Fanuc KAREL source: KX00016.KL

PROGRAM KX00016
%NOLOCKGROUP
VAR
  I: INTEGER
  J: INTEGER
  B: BOOLEAN
  F: FILE
  S: STRING[80]
  P: XYZWPR
BEGIN
  ENABLE CONDITION[1]
END KX00016
